// TIA Portal V21 export
// export: Created 2026-08-21T20:18:56.5598608Z, ExportSetting None, DisplayName Totally Integrated Automation Portal, DisplayVersion V21, DisplayName STEP 7 Professional, DisplayVersion V21, DisplayName STEP 7 Safety, DisplayVersion V21, DisplayName Tech WebApplication, DisplayVersion V21, DisplayName WinCC Basic/Comfort/Advanced, DisplayVersion V21, DisplayName WinCC Professional, DisplayVersion V21, DisplayName WinCC Unified, DisplayVersion V21
TYPE "UDT_Service_Information"
   STRUCT
      state { ExternalWritable := 'False'} : DWord;   // S88 State
      lastState { ExternalWritable := 'False'} : DWord;   // S88 last State
      readyToComplete { ExternalWritable := 'False'} : Bool;   // Ready to complete active
      startTime { ExternalWritable := 'False'} : DTL;   // Start time of control sequence
      endTime { ExternalWritable := 'False'} : DTL;   // End time of control sequence
   END_STRUCT;
END_TYPE
